(* IEC 61131-3 sources: STAR-PLC-Agent/results/raw/four_group_20261114/star_terra/PUB015/generation/sim_00, 1 file *)

(* ---- test_program.st ---- *)
PROGRAM PLC_PRG
VAR
 BenchStep : UDINT := 0;
 BenchCalls : UDINT := 0;
 BenchDone : BOOL := FALSE;
 BenchUut0 : FB_Task;
 BenchUut1 : FB_Task;
 TraceIn_estop : ARRAY[0..15] OF BOOL;
 TraceIn_opeMode : ARRAY[0..15] OF BOOL;
 TraceIn_valveAStart : ARRAY[0..15] OF BOOL;
 TraceIn_valveBStart : ARRAY[0..15] OF BOOL;
 TraceIn_valveCStart : ARRAY[0..15] OF BOOL;
 TraceIn_valveDStart : ARRAY[0..15] OF BOOL;
 TraceIn_mixMotorStart : ARRAY[0..15] OF BOOL;
 TraceIn_autoStart : ARRAY[0..15] OF BOOL;
 TraceIn_processMode : ARRAY[0..15] OF BOOL;
 TraceIn_levelSensor : ARRAY[0..15] OF INT;
 TraceIn_mixMotorComplete : ARRAY[0..15] OF BOOL;
 TraceOut_valveARun : ARRAY[0..15] OF BOOL;
 TraceOut_valveBRun : ARRAY[0..15] OF BOOL;
 TraceOut_valveCRun : ARRAY[0..15] OF BOOL;
 TraceOut_valveDRun : ARRAY[0..15] OF BOOL;
 TraceOut_mixMotorRun : ARRAY[0..15] OF BOOL;
END_VAR

IF NOT BenchDone THEN
 CASE BenchStep OF
 0:
   BenchUut0.estop := TRUE;
   BenchUut0.opeMode := TRUE;
   BenchUut0.valveAStart := FALSE;
   BenchUut0.valveBStart := FALSE;
   BenchUut0.valveCStart := FALSE;
   BenchUut0.valveDStart := FALSE;
   BenchUut0.mixMotorStart := FALSE;
   BenchUut0.autoStart := FALSE;
   BenchUut0.processMode := TRUE;
   BenchUut0.levelSensor := INT#0;
   BenchUut0.mixMotorComplete := FALSE;
   TraceIn_estop[0] := BenchUut0.estop;
   TraceIn_opeMode[0] := BenchUut0.opeMode;
   TraceIn_valveAStart[0] := BenchUut0.valveAStart;
   TraceIn_valveBStart[0] := BenchUut0.valveBStart;
   TraceIn_valveCStart[0] := BenchUut0.valveCStart;
   TraceIn_valveDStart[0] := BenchUut0.valveDStart;
   TraceIn_mixMotorStart[0] := BenchUut0.mixMotorStart;
   TraceIn_autoStart[0] := BenchUut0.autoStart;
   TraceIn_processMode[0] := BenchUut0.processMode;
   TraceIn_levelSensor[0] := BenchUut0.levelSensor;
   TraceIn_mixMotorComplete[0] := BenchUut0.mixMotorComplete;
   BenchUut0();
   TraceOut_valveARun[0] := BenchUut0.valveARun;
   TraceOut_valveBRun[0] := BenchUut0.valveBRun;
   TraceOut_valveCRun[0] := BenchUut0.valveCRun;
   TraceOut_valveDRun[0] := BenchUut0.valveDRun;
   TraceOut_mixMotorRun[0] := BenchUut0.mixMotorRun;
   BenchCalls := BenchCalls + 1;
 1:
   BenchUut0.estop := TRUE;
   BenchUut0.opeMode := TRUE;
   BenchUut0.valveAStart := FALSE;
   BenchUut0.valveBStart := FALSE;
   BenchUut0.valveCStart := FALSE;
   BenchUut0.valveDStart := FALSE;
   BenchUut0.mixMotorStart := FALSE;
   BenchUut0.autoStart := TRUE;
   BenchUut0.processMode := TRUE;
   BenchUut0.levelSensor := INT#49;
   BenchUut0.mixMotorComplete := FALSE;
   TraceIn_estop[1] := BenchUut0.estop;
   TraceIn_opeMode[1] := BenchUut0.opeMode;
   TraceIn_valveAStart[1] := BenchUut0.valveAStart;
   TraceIn_valveBStart[1] := BenchUut0.valveBStart;
   TraceIn_valveCStart[1] := BenchUut0.valveCStart;
   TraceIn_valveDStart[1] := BenchUut0.valveDStart;
   TraceIn_mixMotorStart[1] := BenchUut0.mixMotorStart;
   TraceIn_autoStart[1] := BenchUut0.autoStart;
   TraceIn_processMode[1] := BenchUut0.processMode;
   TraceIn_levelSensor[1] := BenchUut0.levelSensor;
   TraceIn_mixMotorComplete[1] := BenchUut0.mixMotorComplete;
   BenchUut0();
   TraceOut_valveARun[1] := BenchUut0.valveARun;
   TraceOut_valveBRun[1] := BenchUut0.valveBRun;
   TraceOut_valveCRun[1] := BenchUut0.valveCRun;
   TraceOut_valveDRun[1] := BenchUut0.valveDRun;
   TraceOut_mixMotorRun[1] := BenchUut0.mixMotorRun;
   BenchCalls := BenchCalls + 1;
 2:
   BenchUut0.estop := TRUE;
   BenchUut0.opeMode := TRUE;
   BenchUut0.valveAStart := FALSE;
   BenchUut0.valveBStart := FALSE;
   BenchUut0.valveCStart := FALSE;
   BenchUut0.valveDStart := FALSE;
   BenchUut0.mixMotorStart := FALSE;
   BenchUut0.autoStart := FALSE;
   BenchUut0.processMode := FALSE;
   BenchUut0.levelSensor := INT#50;
   BenchUut0.mixMotorComplete := FALSE;
   TraceIn_estop[2] := BenchUut0.estop;
   TraceIn_opeMode[2] := BenchUut0.opeMode;
   TraceIn_valveAStart[2] := BenchUut0.valveAStart;
   TraceIn_valveBStart[2] := BenchUut0.valveBStart;
   TraceIn_valveCStart[2] := BenchUut0.valveCStart;
   TraceIn_valveDStart[2] := BenchUut0.valveDStart;
   TraceIn_mixMotorStart[2] := BenchUut0.mixMotorStart;
   TraceIn_autoStart[2] := BenchUut0.autoStart;
   TraceIn_processMode[2] := BenchUut0.processMode;
   TraceIn_levelSensor[2] := BenchUut0.levelSensor;
   TraceIn_mixMotorComplete[2] := BenchUut0.mixMotorComplete;
   BenchUut0();
   TraceOut_valveARun[2] := BenchUut0.valveARun;
   TraceOut_valveBRun[2] := BenchUut0.valveBRun;
   TraceOut_valveCRun[2] := BenchUut0.valveCRun;
   TraceOut_valveDRun[2] := BenchUut0.valveDRun;
   TraceOut_mixMotorRun[2] := BenchUut0.mixMotorRun;
   BenchCalls := BenchCalls + 1;
 3:
   BenchUut0.estop := TRUE;
   BenchUut0.opeMode := TRUE;
   BenchUut0.valveAStart := FALSE;
   BenchUut0.valveBStart := FALSE;
   BenchUut0.valveCStart := FALSE;
   BenchUut0.valveDStart := FALSE;
   BenchUut0.mixMotorStart := FALSE;
   BenchUut0.autoStart := FALSE;
   BenchUut0.processMode := FALSE;
   BenchUut0.levelSensor := INT#79;
   BenchUut0.mixMotorComplete := FALSE;
   TraceIn_estop[3] := BenchUut0.estop;
   TraceIn_opeMode[3] := BenchUut0.opeMode;
   TraceIn_valveAStart[3] := BenchUut0.valveAStart;
   TraceIn_valveBStart[3] := BenchUut0.valveBStart;
   TraceIn_valveCStart[3] := BenchUut0.valveCStart;
   TraceIn_valveDStart[3] := BenchUut0.valveDStart;
   TraceIn_mixMotorStart[3] := BenchUut0.mixMotorStart;
   TraceIn_autoStart[3] := BenchUut0.autoStart;
   TraceIn_processMode[3] := BenchUut0.processMode;
   TraceIn_levelSensor[3] := BenchUut0.levelSensor;
   TraceIn_mixMotorComplete[3] := BenchUut0.mixMotorComplete;
   BenchUut0();
   TraceOut_valveARun[3] := BenchUut0.valveARun;
   TraceOut_valveBRun[3] := BenchUut0.valveBRun;
   TraceOut_valveCRun[3] := BenchUut0.valveCRun;
   TraceOut_valveDRun[3] := BenchUut0.valveDRun;
   TraceOut_mixMotorRun[3] := BenchUut0.mixMotorRun;
   BenchCalls := BenchCalls + 1;
 4:
   BenchUut0.estop := TRUE;
   BenchUut0.opeMode := TRUE;
   BenchUut0.valveAStart := FALSE;
   BenchUut0.valveBStart := FALSE;
   BenchUut0.valveCStart := FALSE;
   BenchUut0.valveDStart := FALSE;
   BenchUut0.mixMotorStart := FALSE;
   BenchUut0.autoStart := FALSE;
   BenchUut0.processMode := FALSE;
   BenchUut0.levelSensor := INT#80;
   BenchUut0.mixMotorComplete := FALSE;
   TraceIn_estop[4] := BenchUut0.estop;
   TraceIn_opeMode[4] := BenchUut0.opeMode;
   TraceIn_valveAStart[4] := BenchUut0.valveAStart;
   TraceIn_valveBStart[4] := BenchUut0.valveBStart;
   TraceIn_valveCStart[4] := BenchUut0.valveCStart;
   TraceIn_valveDStart[4] := BenchUut0.valveDStart;
   TraceIn_mixMotorStart[4] := BenchUut0.mixMotorStart;
   TraceIn_autoStart[4] := BenchUut0.autoStart;
   TraceIn_processMode[4] := BenchUut0.processMode;
   TraceIn_levelSensor[4] := BenchUut0.levelSensor;
   TraceIn_mixMotorComplete[4] := BenchUut0.mixMotorComplete;
   BenchUut0();
   TraceOut_valveARun[4] := BenchUut0.valveARun;
   TraceOut_valveBRun[4] := BenchUut0.valveBRun;
   TraceOut_valveCRun[4] := BenchUut0.valveCRun;
   TraceOut_valveDRun[4] := BenchUut0.valveDRun;
   TraceOut_mixMotorRun[4] := BenchUut0.mixMotorRun;
   BenchCalls := BenchCalls + 1;
 5:
   BenchUut0.estop := TRUE;
   BenchUut0.opeMode := TRUE;
   BenchUut0.valveAStart := FALSE;
   BenchUut0.valveBStart := FALSE;
   BenchUut0.valveCStart := FALSE;
   BenchUut0.valveDStart := FALSE;
   BenchUut0.mixMotorStart := FALSE;
   BenchUut0.autoStart := FALSE;
   BenchUut0.processMode := FALSE;
   BenchUut0.levelSensor := INT#99;
   BenchUut0.mixMotorComplete := FALSE;
   TraceIn_estop[5] := BenchUut0.estop;
   TraceIn_opeMode[5] := BenchUut0.opeMode;
   TraceIn_valveAStart[5] := BenchUut0.valveAStart;
   TraceIn_valveBStart[5] := BenchUut0.valveBStart;
   TraceIn_valveCStart[5] := BenchUut0.valveCStart;
   TraceIn_valveDStart[5] := BenchUut0.valveDStart;
   TraceIn_mixMotorStart[5] := BenchUut0.mixMotorStart;
   TraceIn_autoStart[5] := BenchUut0.autoStart;
   TraceIn_processMode[5] := BenchUut0.processMode;
   TraceIn_levelSensor[5] := BenchUut0.levelSensor;
   TraceIn_mixMotorComplete[5] := BenchUut0.mixMotorComplete;
   BenchUut0();
   TraceOut_valveARun[5] := BenchUut0.valveARun;
   TraceOut_valveBRun[5] := BenchUut0.valveBRun;
   TraceOut_valveCRun[5] := BenchUut0.valveCRun;
   TraceOut_valveDRun[5] := BenchUut0.valveDRun;
   TraceOut_mixMotorRun[5] := BenchUut0.mixMotorRun;
   BenchCalls := BenchCalls + 1;
 6:
   BenchUut0.estop := TRUE;
   BenchUut0.opeMode := TRUE;
   BenchUut0.valveAStart := FALSE;
   BenchUut0.valveBStart := FALSE;
   BenchUut0.valveCStart := FALSE;
   BenchUut0.valveDStart := FALSE;
   BenchUut0.mixMotorStart := FALSE;
   BenchUut0.autoStart := FALSE;
   BenchUut0.processMode := FALSE;
   BenchUut0.levelSensor := INT#100;
   BenchUut0.mixMotorComplete := FALSE;
   TraceIn_estop[6] := BenchUut0.estop;
   TraceIn_opeMode[6] := BenchUut0.opeMode;
   TraceIn_valveAStart[6] := BenchUut0.valveAStart;
   TraceIn_valveBStart[6] := BenchUut0.valveBStart;
   TraceIn_valveCStart[6] := BenchUut0.valveCStart;
   TraceIn_valveDStart[6] := BenchUut0.valveDStart;
   TraceIn_mixMotorStart[6] := BenchUut0.mixMotorStart;
   TraceIn_autoStart[6] := BenchUut0.autoStart;
   TraceIn_processMode[6] := BenchUut0.processMode;
   TraceIn_levelSensor[6] := BenchUut0.levelSensor;
   TraceIn_mixMotorComplete[6] := BenchUut0.mixMotorComplete;
   BenchUut0();
   TraceOut_valveARun[6] := BenchUut0.valveARun;
   TraceOut_valveBRun[6] := BenchUut0.valveBRun;
   TraceOut_valveCRun[6] := BenchUut0.valveCRun;
   TraceOut_valveDRun[6] := BenchUut0.valveDRun;
   TraceOut_mixMotorRun[6] := BenchUut0.mixMotorRun;
   BenchCalls := BenchCalls + 1;
 7:
   BenchUut0.estop := TRUE;
   BenchUut0.opeMode := TRUE;
   BenchUut0.valveAStart := FALSE;
   BenchUut0.valveBStart := FALSE;
   BenchUut0.valveCStart := FALSE;
   BenchUut0.valveDStart := FALSE;
   BenchUut0.mixMotorStart := FALSE;
   BenchUut0.autoStart := FALSE;
   BenchUut0.processMode := FALSE;
   BenchUut0.levelSensor := INT#100;
   BenchUut0.mixMotorComplete := TRUE;
   TraceIn_estop[7] := BenchUut0.estop;
   TraceIn_opeMode[7] := BenchUut0.opeMode;
   TraceIn_valveAStart[7] := BenchUut0.valveAStart;
   TraceIn_valveBStart[7] := BenchUut0.valveBStart;
   TraceIn_valveCStart[7] := BenchUut0.valveCStart;
   TraceIn_valveDStart[7] := BenchUut0.valveDStart;
   TraceIn_mixMotorStart[7] := BenchUut0.mixMotorStart;
   TraceIn_autoStart[7] := BenchUut0.autoStart;
   TraceIn_processMode[7] := BenchUut0.processMode;
   TraceIn_levelSensor[7] := BenchUut0.levelSensor;
   TraceIn_mixMotorComplete[7] := BenchUut0.mixMotorComplete;
   BenchUut0();
   TraceOut_valveARun[7] := BenchUut0.valveARun;
   TraceOut_valveBRun[7] := BenchUut0.valveBRun;
   TraceOut_valveCRun[7] := BenchUut0.valveCRun;
   TraceOut_valveDRun[7] := BenchUut0.valveDRun;
   TraceOut_mixMotorRun[7] := BenchUut0.mixMotorRun;
   BenchCalls := BenchCalls + 1;
 8:
   BenchUut1.estop := TRUE;
   BenchUut1.opeMode := TRUE;
   BenchUut1.valveAStart := FALSE;
   BenchUut1.valveBStart := FALSE;
   BenchUut1.valveCStart := FALSE;
   BenchUut1.valveDStart := FALSE;
   BenchUut1.mixMotorStart := FALSE;
   BenchUut1.autoStart := FALSE;
   BenchUut1.processMode := FALSE;
   BenchUut1.levelSensor := INT#0;
   BenchUut1.mixMotorComplete := FALSE;
   TraceIn_estop[8] := BenchUut1.estop;
   TraceIn_opeMode[8] := BenchUut1.opeMode;
   TraceIn_valveAStart[8] := BenchUut1.valveAStart;
   TraceIn_valveBStart[8] := BenchUut1.valveBStart;
   TraceIn_valveCStart[8] := BenchUut1.valveCStart;
   TraceIn_valveDStart[8] := BenchUut1.valveDStart;
   TraceIn_mixMotorStart[8] := BenchUut1.mixMotorStart;
   TraceIn_autoStart[8] := BenchUut1.autoStart;
   TraceIn_processMode[8] := BenchUut1.processMode;
   TraceIn_levelSensor[8] := BenchUut1.levelSensor;
   TraceIn_mixMotorComplete[8] := BenchUut1.mixMotorComplete;
   BenchUut1();
   TraceOut_valveARun[8] := BenchUut1.valveARun;
   TraceOut_valveBRun[8] := BenchUut1.valveBRun;
   TraceOut_valveCRun[8] := BenchUut1.valveCRun;
   TraceOut_valveDRun[8] := BenchUut1.valveDRun;
   TraceOut_mixMotorRun[8] := BenchUut1.mixMotorRun;
   BenchCalls := BenchCalls + 1;
 9:
   BenchUut1.estop := TRUE;
   BenchUut1.opeMode := TRUE;
   BenchUut1.valveAStart := FALSE;
   BenchUut1.valveBStart := FALSE;
   BenchUut1.valveCStart := FALSE;
   BenchUut1.valveDStart := FALSE;
   BenchUut1.mixMotorStart := FALSE;
   BenchUut1.autoStart := TRUE;
   BenchUut1.processMode := FALSE;
   BenchUut1.levelSensor := INT#0;
   BenchUut1.mixMotorComplete := FALSE;
   TraceIn_estop[9] := BenchUut1.estop;
   TraceIn_opeMode[9] := BenchUut1.opeMode;
   TraceIn_valveAStart[9] := BenchUut1.valveAStart;
   TraceIn_valveBStart[9] := BenchUut1.valveBStart;
   TraceIn_valveCStart[9] := BenchUut1.valveCStart;
   TraceIn_valveDStart[9] := BenchUut1.valveDStart;
   TraceIn_mixMotorStart[9] := BenchUut1.mixMotorStart;
   TraceIn_autoStart[9] := BenchUut1.autoStart;
   TraceIn_processMode[9] := BenchUut1.processMode;
   TraceIn_levelSensor[9] := BenchUut1.levelSensor;
   TraceIn_mixMotorComplete[9] := BenchUut1.mixMotorComplete;
   BenchUut1();
   TraceOut_valveARun[9] := BenchUut1.valveARun;
   TraceOut_valveBRun[9] := BenchUut1.valveBRun;
   TraceOut_valveCRun[9] := BenchUut1.valveCRun;
   TraceOut_valveDRun[9] := BenchUut1.valveDRun;
   TraceOut_mixMotorRun[9] := BenchUut1.mixMotorRun;
   BenchCalls := BenchCalls + 1;
 10:
   BenchUut1.estop := TRUE;
   BenchUut1.opeMode := TRUE;
   BenchUut1.valveAStart := FALSE;
   BenchUut1.valveBStart := FALSE;
   BenchUut1.valveCStart := FALSE;
   BenchUut1.valveDStart := FALSE;
   BenchUut1.mixMotorStart := FALSE;
   BenchUut1.autoStart := FALSE;
   BenchUut1.processMode := TRUE;
   BenchUut1.levelSensor := INT#51;
   BenchUut1.mixMotorComplete := FALSE;
   TraceIn_estop[10] := BenchUut1.estop;
   TraceIn_opeMode[10] := BenchUut1.opeMode;
   TraceIn_valveAStart[10] := BenchUut1.valveAStart;
   TraceIn_valveBStart[10] := BenchUut1.valveBStart;
   TraceIn_valveCStart[10] := BenchUut1.valveCStart;
   TraceIn_valveDStart[10] := BenchUut1.valveDStart;
   TraceIn_mixMotorStart[10] := BenchUut1.mixMotorStart;
   TraceIn_autoStart[10] := BenchUut1.autoStart;
   TraceIn_processMode[10] := BenchUut1.processMode;
   TraceIn_levelSensor[10] := BenchUut1.levelSensor;
   TraceIn_mixMotorComplete[10] := BenchUut1.mixMotorComplete;
   BenchUut1();
   TraceOut_valveARun[10] := BenchUut1.valveARun;
   TraceOut_valveBRun[10] := BenchUut1.valveBRun;
   TraceOut_valveCRun[10] := BenchUut1.valveCRun;
   TraceOut_valveDRun[10] := BenchUut1.valveDRun;
   TraceOut_mixMotorRun[10] := BenchUut1.mixMotorRun;
   BenchCalls := BenchCalls + 1;
 11:
   BenchUut1.estop := TRUE;
   BenchUut1.opeMode := TRUE;
   BenchUut1.valveAStart := FALSE;
   BenchUut1.valveBStart := FALSE;
   BenchUut1.valveCStart := FALSE;
   BenchUut1.valveDStart := FALSE;
   BenchUut1.mixMotorStart := FALSE;
   BenchUut1.autoStart := FALSE;
   BenchUut1.processMode := TRUE;
   BenchUut1.levelSensor := INT#81;
   BenchUut1.mixMotorComplete := FALSE;
   TraceIn_estop[11] := BenchUut1.estop;
   TraceIn_opeMode[11] := BenchUut1.opeMode;
   TraceIn_valveAStart[11] := BenchUut1.valveAStart;
   TraceIn_valveBStart[11] := BenchUut1.valveBStart;
   TraceIn_valveCStart[11] := BenchUut1.valveCStart;
   TraceIn_valveDStart[11] := BenchUut1.valveDStart;
   TraceIn_mixMotorStart[11] := BenchUut1.mixMotorStart;
   TraceIn_autoStart[11] := BenchUut1.autoStart;
   TraceIn_processMode[11] := BenchUut1.processMode;
   TraceIn_levelSensor[11] := BenchUut1.levelSensor;
   TraceIn_mixMotorComplete[11] := BenchUut1.mixMotorComplete;
   BenchUut1();
   TraceOut_valveARun[11] := BenchUut1.valveARun;
   TraceOut_valveBRun[11] := BenchUut1.valveBRun;
   TraceOut_valveCRun[11] := BenchUut1.valveCRun;
   TraceOut_valveDRun[11] := BenchUut1.valveDRun;
   TraceOut_mixMotorRun[11] := BenchUut1.mixMotorRun;
   BenchCalls := BenchCalls + 1;
 12:
   BenchUut1.estop := FALSE;
   BenchUut1.opeMode := TRUE;
   BenchUut1.valveAStart := FALSE;
   BenchUut1.valveBStart := FALSE;
   BenchUut1.valveCStart := FALSE;
   BenchUut1.valveDStart := FALSE;
   BenchUut1.mixMotorStart := FALSE;
   BenchUut1.autoStart := TRUE;
   BenchUut1.processMode := TRUE;
   BenchUut1.levelSensor := INT#81;
   BenchUut1.mixMotorComplete := TRUE;
   TraceIn_estop[12] := BenchUut1.estop;
   TraceIn_opeMode[12] := BenchUut1.opeMode;
   TraceIn_valveAStart[12] := BenchUut1.valveAStart;
   TraceIn_valveBStart[12] := BenchUut1.valveBStart;
   TraceIn_valveCStart[12] := BenchUut1.valveCStart;
   TraceIn_valveDStart[12] := BenchUut1.valveDStart;
   TraceIn_mixMotorStart[12] := BenchUut1.mixMotorStart;
   TraceIn_autoStart[12] := BenchUut1.autoStart;
   TraceIn_processMode[12] := BenchUut1.processMode;
   TraceIn_levelSensor[12] := BenchUut1.levelSensor;
   TraceIn_mixMotorComplete[12] := BenchUut1.mixMotorComplete;
   BenchUut1();
   TraceOut_valveARun[12] := BenchUut1.valveARun;
   TraceOut_valveBRun[12] := BenchUut1.valveBRun;
   TraceOut_valveCRun[12] := BenchUut1.valveCRun;
   TraceOut_valveDRun[12] := BenchUut1.valveDRun;
   TraceOut_mixMotorRun[12] := BenchUut1.mixMotorRun;
   BenchCalls := BenchCalls + 1;
 13:
   BenchUut1.estop := TRUE;
   BenchUut1.opeMode := TRUE;
   BenchUut1.valveAStart := FALSE;
   BenchUut1.valveBStart := FALSE;
   BenchUut1.valveCStart := FALSE;
   BenchUut1.valveDStart := FALSE;
   BenchUut1.mixMotorStart := FALSE;
   BenchUut1.autoStart := TRUE;
   BenchUut1.processMode := TRUE;
   BenchUut1.levelSensor := INT#0;
   BenchUut1.mixMotorComplete := TRUE;
   TraceIn_estop[13] := BenchUut1.estop;
   TraceIn_opeMode[13] := BenchUut1.opeMode;
   TraceIn_valveAStart[13] := BenchUut1.valveAStart;
   TraceIn_valveBStart[13] := BenchUut1.valveBStart;
   TraceIn_valveCStart[13] := BenchUut1.valveCStart;
   TraceIn_valveDStart[13] := BenchUut1.valveDStart;
   TraceIn_mixMotorStart[13] := BenchUut1.mixMotorStart;
   TraceIn_autoStart[13] := BenchUut1.autoStart;
   TraceIn_processMode[13] := BenchUut1.processMode;
   TraceIn_levelSensor[13] := BenchUut1.levelSensor;
   TraceIn_mixMotorComplete[13] := BenchUut1.mixMotorComplete;
   BenchUut1();
   TraceOut_valveARun[13] := BenchUut1.valveARun;
   TraceOut_valveBRun[13] := BenchUut1.valveBRun;
   TraceOut_valveCRun[13] := BenchUut1.valveCRun;
   TraceOut_valveDRun[13] := BenchUut1.valveDRun;
   TraceOut_mixMotorRun[13] := BenchUut1.mixMotorRun;
   BenchCalls := BenchCalls + 1;
 14:
   BenchUut1.estop := TRUE;
   BenchUut1.opeMode := TRUE;
   BenchUut1.valveAStart := FALSE;
   BenchUut1.valveBStart := FALSE;
   BenchUut1.valveCStart := FALSE;
   BenchUut1.valveDStart := FALSE;
   BenchUut1.mixMotorStart := FALSE;
   BenchUut1.autoStart := FALSE;
   BenchUut1.processMode := TRUE;
   BenchUut1.levelSensor := INT#0;
   BenchUut1.mixMotorComplete := FALSE;
   TraceIn_estop[14] := BenchUut1.estop;
   TraceIn_opeMode[14] := BenchUut1.opeMode;
   TraceIn_valveAStart[14] := BenchUut1.valveAStart;
   TraceIn_valveBStart[14] := BenchUut1.valveBStart;
   TraceIn_valveCStart[14] := BenchUut1.valveCStart;
   TraceIn_valveDStart[14] := BenchUut1.valveDStart;
   TraceIn_mixMotorStart[14] := BenchUut1.mixMotorStart;
   TraceIn_autoStart[14] := BenchUut1.autoStart;
   TraceIn_processMode[14] := BenchUut1.processMode;
   TraceIn_levelSensor[14] := BenchUut1.levelSensor;
   TraceIn_mixMotorComplete[14] := BenchUut1.mixMotorComplete;
   BenchUut1();
   TraceOut_valveARun[14] := BenchUut1.valveARun;
   TraceOut_valveBRun[14] := BenchUut1.valveBRun;
   TraceOut_valveCRun[14] := BenchUut1.valveCRun;
   TraceOut_valveDRun[14] := BenchUut1.valveDRun;
   TraceOut_mixMotorRun[14] := BenchUut1.mixMotorRun;
   BenchCalls := BenchCalls + 1;
 15:
   BenchUut1.estop := TRUE;
   BenchUut1.opeMode := TRUE;
   BenchUut1.valveAStart := FALSE;
   BenchUut1.valveBStart := FALSE;
   BenchUut1.valveCStart := FALSE;
   BenchUut1.valveDStart := FALSE;
   BenchUut1.mixMotorStart := FALSE;
   BenchUut1.autoStart := TRUE;
   BenchUut1.processMode := TRUE;
   BenchUut1.levelSensor := INT#0;
   BenchUut1.mixMotorComplete := FALSE;
   TraceIn_estop[15] := BenchUut1.estop;
   TraceIn_opeMode[15] := BenchUut1.opeMode;
   TraceIn_valveAStart[15] := BenchUut1.valveAStart;
   TraceIn_valveBStart[15] := BenchUut1.valveBStart;
   TraceIn_valveCStart[15] := BenchUut1.valveCStart;
   TraceIn_valveDStart[15] := BenchUut1.valveDStart;
   TraceIn_mixMotorStart[15] := BenchUut1.mixMotorStart;
   TraceIn_autoStart[15] := BenchUut1.autoStart;
   TraceIn_processMode[15] := BenchUut1.processMode;
   TraceIn_levelSensor[15] := BenchUut1.levelSensor;
   TraceIn_mixMotorComplete[15] := BenchUut1.mixMotorComplete;
   BenchUut1();
   TraceOut_valveARun[15] := BenchUut1.valveARun;
   TraceOut_valveBRun[15] := BenchUut1.valveBRun;
   TraceOut_valveCRun[15] := BenchUut1.valveCRun;
   TraceOut_valveDRun[15] := BenchUut1.valveDRun;
   TraceOut_mixMotorRun[15] := BenchUut1.mixMotorRun;
   BenchCalls := BenchCalls + 1;
 END_CASE;
 BenchStep := BenchStep + 1;
 IF BenchStep >= 16 THEN BenchDone := TRUE; END_IF;
END_IF;
END_PROGRAM
